// TIA Portal V19 export
// export: Created 2026-11-08T08:30:00.0000000Z, ExportSetting WithReadOnly
DATA_BLOCK "DB_ExampleData"   // DB1
{ S7_Optimized_Access := 'TRUE' }
// stored: IsOnlyStoredInLoadMemory false, IsWriteProtectedInAS false
   VAR
      Speed : Real := 0.0;
      Scaled : Int;
   END_VAR
   VAR RETAIN
      Limit { S7_SetPoint := 'True'} : Real := 90.0;   // High speed limit
   END_VAR
   VAR
      Cfg : Struct
         Enable : Bool := true;
         Delay : Time := T#5S;
      END_STRUCT;
      Steps : Array[0..1] of Int;
   END_VAR
BEGIN
   Steps[0] := 10;
   Steps[1] := 20;
END_DATA_BLOCK
